// Core 10.5.1: identity is fixed at generation; the publisher writes live state.
DATA_BLOCK "GDB_PressDemoFieldbus"
{ S7_Optimized_Access := 'TRUE' }
VERSION : 0.1
NON_RETAIN
VAR
    Topology {ExternalWritable := 'False'} : "ST_FieldbusTopology";
END_VAR
BEGIN
    Topology.NodeCount := 3;
    Topology.MappingValid := TRUE;
    Topology.Nodes[1].Name := 'PressIo1214C';
    Topology.Nodes[1].DescriptionKey := 'project.hardware.s71214c';
    Topology.Nodes[1].TypeId := 'CPU 1214C DC/DC/DC 6ES7 214-1AG40-0XB0';
    Topology.Nodes[1].Address := '192.168.0.10 (I/O bridge)';
    Topology.Nodes[1].ParentIdx := 0;
    Topology.Nodes[1].ChannelCount := 0;
    Topology.Nodes[2].Name := 'PressIo1214C DI';
    Topology.Nodes[2].DescriptionKey := 'project.hardware.s71214cDi';
    Topology.Nodes[2].TypeId := 'Onboard DI 14 x 24 V DC';
    Topology.Nodes[2].Address := '%I0.0..%I1.5';
    Topology.Nodes[2].ParentIdx := 1;
    Topology.Nodes[2].ChannelCount := 14;
    Topology.Nodes[2].Channels[1].Name := '_101B301A';
    Topology.Nodes[2].Channels[1].DescriptionKey := 'project.io.101B301A';
    Topology.Nodes[2].Channels[1].Address := '%I0.0';
    Topology.Nodes[2].Channels[1].Path := WSTRING#'PressIo1214C DI/_101B301A';
    Topology.Nodes[2].Channels[1].ModulePath := WSTRING#'PressDemo.PartSlide';
    Topology.Nodes[2].Channels[1].Dir := 0;
    Topology.Nodes[2].Channels[1].Kind := 0;
    Topology.Nodes[2].Channels[2].Name := '_101B301B';
    Topology.Nodes[2].Channels[2].DescriptionKey := 'project.io.101B301B';
    Topology.Nodes[2].Channels[2].Address := '%I0.1';
    Topology.Nodes[2].Channels[2].Path := WSTRING#'PressIo1214C DI/_101B301B';
    Topology.Nodes[2].Channels[2].ModulePath := WSTRING#'PressDemo.PartSlide';
    Topology.Nodes[2].Channels[2].Dir := 0;
    Topology.Nodes[2].Channels[2].Kind := 0;
    Topology.Nodes[2].Channels[3].Name := '_101B201A';
    Topology.Nodes[2].Channels[3].DescriptionKey := 'project.io.101B201A';
    Topology.Nodes[2].Channels[3].Address := '%I0.2';
    Topology.Nodes[2].Channels[3].Path := WSTRING#'PressIo1214C DI/_101B201A';
    Topology.Nodes[2].Channels[3].ModulePath := WSTRING#'PressDemo.Door';
    Topology.Nodes[2].Channels[3].Dir := 0;
    Topology.Nodes[2].Channels[3].Kind := 0;
    Topology.Nodes[2].Channels[4].Name := '_101B201B';
    Topology.Nodes[2].Channels[4].DescriptionKey := 'project.io.101B201B';
    Topology.Nodes[2].Channels[4].Address := '%I0.3';
    Topology.Nodes[2].Channels[4].Path := WSTRING#'PressIo1214C DI/_101B201B';
    Topology.Nodes[2].Channels[4].ModulePath := WSTRING#'PressDemo.Door';
    Topology.Nodes[2].Channels[4].Dir := 0;
    Topology.Nodes[2].Channels[4].Kind := 0;
    Topology.Nodes[2].Channels[5].Name := '_101B202A';
    Topology.Nodes[2].Channels[5].DescriptionKey := 'project.io.101B202A';
    Topology.Nodes[2].Channels[5].Address := '%I0.4';
    Topology.Nodes[2].Channels[5].Path := WSTRING#'PressIo1214C DI/_101B202A';
    Topology.Nodes[2].Channels[5].ModulePath := WSTRING#'PressDemo.PressRam';
    Topology.Nodes[2].Channels[5].Dir := 0;
    Topology.Nodes[2].Channels[5].Kind := 0;
    Topology.Nodes[2].Channels[6].Name := '_101B202B';
    Topology.Nodes[2].Channels[6].DescriptionKey := 'project.io.101B202B';
    Topology.Nodes[2].Channels[6].Address := '%I0.5';
    Topology.Nodes[2].Channels[6].Path := WSTRING#'PressIo1214C DI/_101B202B';
    Topology.Nodes[2].Channels[6].ModulePath := WSTRING#'PressDemo.PressRam';
    Topology.Nodes[2].Channels[6].Dir := 0;
    Topology.Nodes[2].Channels[6].Kind := 0;
    Topology.Nodes[2].Channels[7].Name := '_101S101';
    Topology.Nodes[2].Channels[7].DescriptionKey := 'project.io.101S101';
    Topology.Nodes[2].Channels[7].Address := '%I0.6';
    Topology.Nodes[2].Channels[7].Path := WSTRING#'PressIo1214C DI/_101S101';
    Topology.Nodes[2].Channels[7].ModulePath := WSTRING#'PressDemo.TwoHand';
    Topology.Nodes[2].Channels[7].Dir := 0;
    Topology.Nodes[2].Channels[7].Kind := 0;
    Topology.Nodes[2].Channels[8].Name := '_101S102';
    Topology.Nodes[2].Channels[8].DescriptionKey := 'project.io.101S102';
    Topology.Nodes[2].Channels[8].Address := '%I0.7';
    Topology.Nodes[2].Channels[8].Path := WSTRING#'PressIo1214C DI/_101S102';
    Topology.Nodes[2].Channels[8].ModulePath := WSTRING#'PressDemo.TwoHand';
    Topology.Nodes[2].Channels[8].Dir := 0;
    Topology.Nodes[2].Channels[8].Kind := 0;
    Topology.Nodes[2].Channels[9].Name := '_000MB085A_2';
    Topology.Nodes[2].Channels[9].DescriptionKey := 'project.io.000MB085A_2';
    Topology.Nodes[2].Channels[9].Address := '%I1.0';
    Topology.Nodes[2].Channels[9].Path := WSTRING#'PressIo1214C DI/_000MB085A_2';
    Topology.Nodes[2].Channels[9].ModulePath := WSTRING#'PressDemo.AirPressureMonitor';
    Topology.Nodes[2].Channels[9].Dir := 0;
    Topology.Nodes[2].Channels[9].Kind := 0;
    Topology.Nodes[2].Channels[10].Name := '_000MB085A_4';
    Topology.Nodes[2].Channels[10].DescriptionKey := 'project.io.000MB085A_4';
    Topology.Nodes[2].Channels[10].Address := '%I1.1';
    Topology.Nodes[2].Channels[10].Path := WSTRING#'PressIo1214C DI/_000MB085A_4';
    Topology.Nodes[2].Channels[10].ModulePath := WSTRING#'PressDemo.AirPressureMonitor';
    Topology.Nodes[2].Channels[10].Dir := 0;
    Topology.Nodes[2].Channels[10].Kind := 0;
    Topology.Nodes[2].Channels[11].Name := '_101B601';
    Topology.Nodes[2].Channels[11].DescriptionKey := 'project.io.101B601';
    Topology.Nodes[2].Channels[11].Address := '%I1.2';
    Topology.Nodes[2].Channels[11].Path := WSTRING#'PressIo1214C DI/_101B601';
    Topology.Nodes[2].Channels[11].ModulePath := WSTRING#'PressDemo.PartPresentSensor';
    Topology.Nodes[2].Channels[11].Dir := 0;
    Topology.Nodes[2].Channels[11].Kind := 0;
    Topology.Nodes[2].Channels[12].Name := '_000K911_Y32';
    Topology.Nodes[2].Channels[12].DescriptionKey := 'project.io.000K911_Y32';
    Topology.Nodes[2].Channels[12].Address := '%I1.3';
    Topology.Nodes[2].Channels[12].Path := WSTRING#'PressIo1214C DI/_000K911_Y32';
    Topology.Nodes[2].Channels[12].ModulePath := WSTRING#'PressDemo';
    Topology.Nodes[2].Channels[12].Dir := 0;
    Topology.Nodes[2].Channels[12].Kind := 0;
    Topology.Nodes[2].Channels[13].Name := '_000K910A';
    Topology.Nodes[2].Channels[13].DescriptionKey := 'project.io.000K910A';
    Topology.Nodes[2].Channels[13].Address := '%I1.4';
    Topology.Nodes[2].Channels[13].Path := WSTRING#'PressIo1214C DI/_000K910A';
    Topology.Nodes[2].Channels[13].ModulePath := WSTRING#'PressDemo';
    Topology.Nodes[2].Channels[13].Dir := 0;
    Topology.Nodes[2].Channels[13].Kind := 0;
    Topology.Nodes[2].Channels[14].Name := '_EvaluatedTwoHand';
    Topology.Nodes[2].Channels[14].DescriptionKey := 'project.io.EvaluatedTwoHand';
    Topology.Nodes[2].Channels[14].Address := '%I1.5';
    Topology.Nodes[2].Channels[14].Path := WSTRING#'PressIo1214C DI/_EvaluatedTwoHand';
    Topology.Nodes[2].Channels[14].ModulePath := WSTRING#'PressDemo.TwoHand';
    Topology.Nodes[2].Channels[14].Dir := 0;
    Topology.Nodes[2].Channels[14].Kind := 0;
    Topology.Nodes[3].Name := 'PressIo1214C DQ';
    Topology.Nodes[3].DescriptionKey := 'project.hardware.s71214cDq';
    Topology.Nodes[3].TypeId := 'Onboard DQ 10 x 24 V DC';
    Topology.Nodes[3].Address := '%Q0.0..%Q1.1';
    Topology.Nodes[3].ParentIdx := 1;
    Topology.Nodes[3].ChannelCount := 10;
    Topology.Nodes[3].Channels[1].Name := '_101K301A';
    Topology.Nodes[3].Channels[1].DescriptionKey := 'project.io.101K301A';
    Topology.Nodes[3].Channels[1].Address := '%Q0.0';
    Topology.Nodes[3].Channels[1].Path := WSTRING#'PressIo1214C DQ/_101K301A';
    Topology.Nodes[3].Channels[1].ModulePath := WSTRING#'PressDemo.PartSlide';
    Topology.Nodes[3].Channels[1].Dir := 1;
    Topology.Nodes[3].Channels[1].Kind := 0;
    Topology.Nodes[3].Channels[2].Name := '_101K301B';
    Topology.Nodes[3].Channels[2].DescriptionKey := 'project.io.101K301B';
    Topology.Nodes[3].Channels[2].Address := '%Q0.1';
    Topology.Nodes[3].Channels[2].Path := WSTRING#'PressIo1214C DQ/_101K301B';
    Topology.Nodes[3].Channels[2].ModulePath := WSTRING#'PressDemo.PartSlide';
    Topology.Nodes[3].Channels[2].Dir := 1;
    Topology.Nodes[3].Channels[2].Kind := 0;
    Topology.Nodes[3].Channels[3].Name := '_101K201A';
    Topology.Nodes[3].Channels[3].DescriptionKey := 'project.io.101K201A';
    Topology.Nodes[3].Channels[3].Address := '%Q0.2';
    Topology.Nodes[3].Channels[3].Path := WSTRING#'PressIo1214C DQ/_101K201A';
    Topology.Nodes[3].Channels[3].ModulePath := WSTRING#'PressDemo.Door';
    Topology.Nodes[3].Channels[3].Dir := 1;
    Topology.Nodes[3].Channels[3].Kind := 0;
    Topology.Nodes[3].Channels[4].Name := '_101K201B';
    Topology.Nodes[3].Channels[4].DescriptionKey := 'project.io.101K201B';
    Topology.Nodes[3].Channels[4].Address := '%Q0.3';
    Topology.Nodes[3].Channels[4].Path := WSTRING#'PressIo1214C DQ/_101K201B';
    Topology.Nodes[3].Channels[4].ModulePath := WSTRING#'PressDemo.Door';
    Topology.Nodes[3].Channels[4].Dir := 1;
    Topology.Nodes[3].Channels[4].Kind := 0;
    Topology.Nodes[3].Channels[5].Name := '_101K202A';
    Topology.Nodes[3].Channels[5].DescriptionKey := 'project.io.101K202A';
    Topology.Nodes[3].Channels[5].Address := '%Q0.4';
    Topology.Nodes[3].Channels[5].Path := WSTRING#'PressIo1214C DQ/_101K202A';
    Topology.Nodes[3].Channels[5].ModulePath := WSTRING#'PressDemo.PressRam';
    Topology.Nodes[3].Channels[5].Dir := 1;
    Topology.Nodes[3].Channels[5].Kind := 0;
    Topology.Nodes[3].Channels[6].Name := '_101K202B';
    Topology.Nodes[3].Channels[6].DescriptionKey := 'project.io.101K202B';
    Topology.Nodes[3].Channels[6].Address := '%Q0.5';
    Topology.Nodes[3].Channels[6].Path := WSTRING#'PressIo1214C DQ/_101K202B';
    Topology.Nodes[3].Channels[6].ModulePath := WSTRING#'PressDemo.PressRam';
    Topology.Nodes[3].Channels[6].Dir := 1;
    Topology.Nodes[3].Channels[6].Kind := 0;
    Topology.Nodes[3].Channels[7].Name := '_101P101';
    Topology.Nodes[3].Channels[7].DescriptionKey := 'project.io.101P101';
    Topology.Nodes[3].Channels[7].Address := '%Q0.6';
    Topology.Nodes[3].Channels[7].Path := WSTRING#'PressIo1214C DQ/_101P101';
    Topology.Nodes[3].Channels[7].ModulePath := WSTRING#'PressDemo';
    Topology.Nodes[3].Channels[7].Dir := 1;
    Topology.Nodes[3].Channels[7].Kind := 0;
    Topology.Nodes[3].Channels[8].Name := '_101P102';
    Topology.Nodes[3].Channels[8].DescriptionKey := 'project.io.101P102';
    Topology.Nodes[3].Channels[8].Address := '%Q0.7';
    Topology.Nodes[3].Channels[8].Path := WSTRING#'PressIo1214C DQ/_101P102';
    Topology.Nodes[3].Channels[8].ModulePath := WSTRING#'PressDemo';
    Topology.Nodes[3].Channels[8].Dir := 1;
    Topology.Nodes[3].Channels[8].Kind := 0;
    Topology.Nodes[3].Channels[9].Name := '_000K951_A1';
    Topology.Nodes[3].Channels[9].DescriptionKey := 'project.io.000K951_A1';
    Topology.Nodes[3].Channels[9].Address := '%Q1.0';
    Topology.Nodes[3].Channels[9].Path := WSTRING#'PressIo1214C DQ/_000K951_A1';
    Topology.Nodes[3].Channels[9].ModulePath := WSTRING#'PressDemo';
    Topology.Nodes[3].Channels[9].Dir := 1;
    Topology.Nodes[3].Channels[9].Kind := 0;
    Topology.Nodes[3].Channels[10].Name := '_000K911_A1';
    Topology.Nodes[3].Channels[10].DescriptionKey := 'project.io.000K911_A1';
    Topology.Nodes[3].Channels[10].Address := '%Q1.1';
    Topology.Nodes[3].Channels[10].Path := WSTRING#'PressIo1214C DQ/_000K911_A1';
    Topology.Nodes[3].Channels[10].ModulePath := WSTRING#'PressDemo';
    Topology.Nodes[3].Channels[10].Dir := 1;
    Topology.Nodes[3].Channels[10].Kind := 0;
END_DATA_BLOCK
